TYPE ST_ITECH_SetConfigs :
STRUCT
	dcSource	: ST_ITECH_DCSource;
	protection	: ST_ITECH_Protection;
END_STRUCT
END_TYPE

(* stored: Version 1.1.0.1
   DUT ST_ITECH_SetConfigs: Id {e199adfe-3f29-431f-8931-081e040dc22c} *)
